(* IEC 61131-3 sources: guidance-for-physical-ai-production-designer-on-aws/source/plan2cell/crates/bt2plc/tests/golden/cell_2robot/codesys/robots/robot1/GVL, 1 file *)

(* ---- GVL_Program.st ---- *)
(*
 * GVL_Program - generated by bt2plc 0.1.0 - DO NOT EDIT
 * Robot program of robot1 (R1) for plan bt_1791274820_cell_2robot (cell cell_2robot)
 * Angles in degrees (KUKA A1..A6 after joint sign/offset), times in seconds from op start.
 *)
{attribute 'qualified_only'}
VAR_GLOBAL CONSTANT
    (* ========================================================================
       IDENTITY / PROTOCOL
       ======================================================================== *)
    ROBOT_TAG               : STRING(16) := 'R1';
    ROBOT_NS                : STRING(32) := 'robot1';
    ROBOT_INDEX             : WORD := WORD#1;
    PLAN_ID                 : WORD := WORD#16#A312;             (* must match the head PLC *)
    PROD_FOLGE              : WORD := WORD#11;
    HOME_FOLGE              : WORD := WORD#125;
    JOB_NUMBER_BYTE         : BOOL := FALSE;
    STEP_BYTE               : INT := 4;
    REQ_BYTE                : INT := 28;
    GRANT_BYTE              : INT := 12;
    PLAN_ID_BYTE            : INT := 4;
    R_TASK_S                : REAL := 0.0200;                   (* device MainTask interval *)
    R_HOME_S                : REAL := 7.0000;                   (* blind home duration *)
    R_AT_HOME_TOL_DEG       : REAL := 0.5000;
    R_START_TOL_DEG         : REAL := 1.0000;
    ERR_UNKNOWN_FOLGE       : WORD := WORD#16#0101;
    ERR_PLAN_MISMATCH       : WORD := WORD#16#0103;
    WARN_START_DEVIATION    : WORD := WORD#16#0201;

    (* ========================================================================
       PROGRAM
       ======================================================================== *)
    N_OPS                   : INT := 2;
    N_WP                    : INT := 27;
    arHomeDeg               : ARRAY[1..6] OF REAL := [0.0000, -90.0000, 90.0000, 0.0000, 0.0000, 0.0000];
    aOps                    : ARRAY[1..2] OF ST_OpDef := [
        (sName := 'STAGE_R1', nFirstWp := 1, nLastWp := 14, dwZoneMask := DWORD#16#00000000, tDelay := T#0MS, tHold := T#500MS, rDelay_s := 0.0000, rHold_s := 0.5000, rVelScale := 1.0000, bBlindHome := FALSE),    (* #1 STAGE_R1 (move) *)
        (sName := 'HOME', nFirstWp := 15, nLastWp := 27, dwZoneMask := DWORD#16#00000000, tDelay := T#0MS, tHold := T#0MS, rDelay_s := 0.0000, rHold_s := 0.0000, rVelScale := 1.0000, bBlindHome := FALSE)    (* #2 HOME (home) *)
    ];
    aWp                     : ARRAY[1..27] OF ST_Waypoint := [
        (* op 1 STAGE_R1 - traj_robot1_STAGE_R1 *)
        (rT := 0.0000, rA1 := 0.0000, rA2 := -90.0000, rA3 := 90.0000, rA4 := 0.0000, rA5 := 0.0000, rA6 := 0.0000),
        (rT := 0.2767, rA1 := 0.1421, rA2 := -89.0006, rA3 := 89.9771, rA4 := 0.0000, rA5 := 0.0000, rA6 := 0.0000),
        (rT := 0.5530, rA1 := 0.5354, rA2 := -86.2310, rA3 := 89.9133, rA4 := 0.0000, rA5 := 0.0000, rA6 := 0.0000),
        (rT := 0.8297, rA1 := 1.1310, rA2 := -82.0342, rA3 := 89.8161, rA4 := 0.0000, rA5 := 0.0000, rA6 := 0.0000),
        (rT := 1.1063, rA1 := 1.8795, rA2 := -76.7531, rA3 := 89.6931, rA4 := 0.0000, rA5 := 0.0000, rA6 := 0.0000),
        (rT := 1.3830, rA1 := 2.7319, rA2 := -70.7305, rA3 := 89.5515, rA4 := 0.0000, rA5 := 0.0000, rA6 := 0.0000),
        (rT := 1.6593, rA1 := 3.6388, rA2 := -64.3095, rA3 := 89.3990, rA4 := 0.0000, rA5 := 0.0000, rA6 := 0.0000),
        (rT := 1.9360, rA1 := 4.5513, rA2 := -57.8329, rA3 := 89.2429, rA4 := 0.0000, rA5 := 0.0000, rA6 := 0.0000),
        (rT := 2.2127, rA1 := 5.4200, rA2 := -51.6436, rA3 := 89.0908, rA4 := 0.0000, rA5 := 0.0000, rA6 := 0.0000),
        (rT := 2.4893, rA1 := 6.1959, rA2 := -46.0847, rA3 := 88.9501, rA4 := 0.0000, rA5 := 0.0000, rA6 := 0.0000),
        (rT := 2.7657, rA1 := 6.8297, rA2 := -41.4990, rA3 := 88.8283, rA4 := 0.0000, rA5 := 0.0000, rA6 := 0.0000),
        (rT := 3.0423, rA1 := 7.2722, rA2 := -38.2294, rA3 := 88.7329, rA4 := 0.0000, rA5 := 0.0000, rA6 := 0.0000),
        (rT := 3.1357, rA1 := 7.7267, rA2 := -33.2119, rA3 := 88.3788, rA4 := 0.0000, rA5 := 0.0000, rA6 := 0.0000),
        (rT := 3.2287, rA1 := 7.2722, rA2 := -35.0616, rA3 := 88.2443, rA4 := 0.0000, rA5 := 0.0000, rA6 := 0.0000),
        (* op 2 HOME - traj_robot1_n3 *)
        (rT := 0.0000, rA1 := 7.2722, rA2 := -35.0616, rA3 := 88.2443, rA4 := 0.0000, rA5 := 0.0000, rA6 := 0.0000),
        (rT := 0.2015, rA1 := 7.1292, rA2 := -36.1426, rA3 := 88.2788, rA4 := 0.0000, rA5 := 0.0000, rA6 := 0.0000),
        (rT := 0.4032, rA1 := 6.7336, rA2 := -39.1311, rA3 := 88.3743, rA4 := 0.0000, rA5 := 0.0000, rA6 := 0.0000),
        (rT := 0.6048, rA1 := 6.1360, rA2 := -43.6457, rA3 := 88.5186, rA4 := 0.0000, rA5 := 0.0000, rA6 := 0.0000),
        (rT := 0.8065, rA1 := 5.3868, rA2 := -49.3049, rA3 := 88.6995, rA4 := 0.0000, rA5 := 0.0000, rA6 := 0.0000),
        (rT := 1.0080, rA1 := 4.5367, rA2 := -55.7271, rA3 := 88.9047, rA4 := 0.0000, rA5 := 0.0000, rA6 := 0.0000),
        (rT := 1.2097, rA1 := 3.6361, rA2 := -62.5308, rA3 := 89.1221, rA4 := 0.0000, rA5 := 0.0000, rA6 := 0.0000),
        (rT := 1.4112, rA1 := 2.7355, rA2 := -69.3345, rA3 := 89.3396, rA4 := 0.0000, rA5 := 0.0000, rA6 := 0.0000),
        (rT := 1.6127, rA1 := 1.8854, rA2 := -75.7567, rA3 := 89.5448, rA4 := 0.0000, rA5 := 0.0000, rA6 := 0.0000),
        (rT := 1.8145, rA1 := 1.1363, rA2 := -81.4159, rA3 := 89.7257, rA4 := 0.0000, rA5 := 0.0000, rA6 := 0.0000),
        (rT := 2.0160, rA1 := 0.5387, rA2 := -85.9305, rA3 := 89.8699, rA4 := 0.0000, rA5 := 0.0000, rA6 := 0.0000),
        (rT := 2.2177, rA1 := 0.1431, rA2 := -88.9190, rA3 := 89.9655, rA4 := 0.0000, rA5 := 0.0000, rA6 := 0.0000),
        (rT := 2.4192, rA1 := 0.0000, rA2 := -90.0000, rA3 := 90.0000, rA4 := 0.0000, rA5 := 0.0000, rA6 := 0.0000)
    ];
END_VAR
